(* IEC 61131-3 sources: SortJet_MasterSPS_Aufbau.fbsproj/07_Auftragsverwaltung/BasisSchrittketten (part 3) *)

(* ---- TS_Eintransport.fb.st ---- *)
(* METADATA
{
	"v3Meta": {
		"objectGuid": "2467a7d0-b543-4c0f-8e2f-d0f3bb8e773e"
	}
}
*)
FUNCTION_BLOCK TS_Eintransport
VAR_INPUT

  // BOOLEAN
  bpReset                : BOOL;

  // WORD
  wStation               : WORD;

  // STRUKTUR
  Auftragsdaten          : Auftragsdaten_ST;

END_VAR
VAR_OUTPUT

  // BOOLEAN
  bpDone                 : BOOL;
  bpFehler               : BOOL;

END_VAR
VAR
  // BOOLEAN
  blStationQuittiertScheiben : BOOL;

  // WORD
  wlEintransportstation  : WORD;

  // INT
  ilScheibenZuQuittieren : INT;

  // STEPS
  steplSchritt           : STEPS_TE;

END_VAR

//-------------------------------------------------------------------------------------------------
// STEUERUNG: EINTRANSPORT
//-------------------------------------------------------------------------------------------------
IF ( Auftragsdaten.wAuftrag = eStation_Eintransport ) THEN
  CASE steplSchritt OF
    // EINTRANSPORT  =============================== ============
    STEP_0_E:
      (* Hinweis:
         - Ueberpruefen des Sicherheitskreises
      *)
      IF  (checkSafetyCircuitsNotBlocked(starrTransferShuttleBasisParameter[wStation])
            AND NOT starrTransfershuttleBasisParameter[wStation].bReset )
      THEN
        steplSchritt := STEP_100_E;
      END_IF

    // EINTRANSPORT  ===========================================
    STEP_100_E:
      (* Anmerkung:
         - Zielstation abfragen ob diese bereit ist zum Austransport
      *)
      wlEintransportstation := Auftragsdaten.wTransferstationsNr1;
      ilScheibenZuQuittieren := WORD_TO_INT( Auftragsdaten.wAnzahlScheiben);

      CASE wlEintransportstation OF

          (* Hinweis:
             - Ruecktransport durch den Speicher beruecksichtigen
          *)
          cERSTES_INPUTSHUTTLE..cLETZTES_INPUTSHUTTLE,
            cERSTES_OUTPUTSHUTTLE..cLETZTES_OUTPUTSHUTTLE:
          IF ( Job_Shuttle.AuftragsdatenWand[Auftragsdaten.wTransferstationsNr1, Auftragsdaten.wTransferwand].wAuftrag = eStation_Austransport ) THEN
            steplSchritt := STEP_110_E;

          ELSE
            wpgFehlerdaten[0] := starrTransfershuttleBasisParameter[wStation].stMKs.stStationsNummern.NummerExtern;
            wpgFehlerdaten[1] := wlEintransportstation;
            wpgFehlerdaten[2] := Job_Shuttle.AuftragsdatenWand[Auftragsdaten.wTransferstationsNr1, Auftragsdaten.wTransferwand].wAuftrag;

            SpsError( eFehler_Station,
                      cMELDUNG_AUFTRAGSDATEN_AUFTRAGSTATUS_GLAS_SENDER_UNGUELTIG,
                      starrTransfershuttleBasisParameter[wStation].stMKs.stStationsNummern.NummerIntern,
                      AutomatikkreisBestimmen(starrTransfershuttleBasisParameter[wStation].stMKs.stStationsNummern.NummerSPS),
                      wpgFehlerdaten );

            steplSchritt := STEP_900_E;
          END_IF

        // Stationen
        //   - Wie beim Shuttle: Der TS legt den Austransport-Auftrag der Station an, sobald sie belegt ist
        cERSTE_STATION..cLETZTE_STATION:
          IF (    ( Job_Stationen.AuftragsdatenWand[wlEintransportstation, Auftragsdaten.wTransferwand].wAuftrag = eStation_Belegt )
               OR ( Job_Stationen.AuftragsdatenWand[wlEintransportstation, Auftragsdaten.wTransferwand].wAuftrag = eStation_Warte_Auf_Austransport ) )
             AND AutomatikAktiv(wlEintransportstation)
          THEN

            Job_Stationen.AuftragsdatenWand[wlEintransportstation, Auftragsdaten.wTransferwand]          := AuftragsdatenUmkopieren(FALSE, FALSE, Auftragsdaten);
            Job_Stationen.AuftragsdatenWand[wlEintransportstation, Auftragsdaten.wTransferwand].wAuftrag := eStation_Austransport;

            // Kopplung zur Station herstellen
            starrTransfershuttleBasisParameter[wStation].InGlasTransportNachfolger[cWAND_1] := starrStationBasisParameter[wlEintransportstation].OutGlasTransport[Auftragsdaten.wTransferwand];
            starrTransfershuttleBasisParameter[wStation].InGlasTransportVorgaenger[cWAND_1] := starrStationBasisParameter[wlEintransportstation].OutGlasTransport[Auftragsdaten.wTransferwand];

            steplSchritt := STEP_110_E;
          END_IF

        ELSE
          wpgFehlerdaten[0] := starrTransfershuttleBasisParameter[wStation].stMKs.stStationsNummern.NummerExtern;
          wpgFehlerdaten[1] := wlEintransportstation;

          SpsError( eFehler_Station,
                    cMELDUNG_AUFTRAGSDATEN_FALSCHE_EINLAUFSTATION,
                    starrTransfershuttleBasisParameter[wStation].stMKs.stStationsNummern.NummerIntern,
                    AutomatikkreisBestimmen(starrTransfershuttleBasisParameter[wStation].stMKs.stStationsNummern.NummerSPS),
                    wpgFehlerdaten );

          steplSchritt := STEP_900_E;

      END_CASE

      (* Fehlerbehandlung:
         - Shuttle
      *)
      IF ( starrTransfershuttleBasisParameter[wStation].bFehler ) THEN

        SpsError( eFehler_Station,
                  starrTransfershuttleBasisParameter[wStation].wFehlerNummer,
                  starrTransfershuttleBasisParameter[wStation].stMKs.stStationsNummern.NummerIntern,
                  AutomatikkreisBestimmen(starrTransfershuttleBasisParameter[wStation].stMKs.stStationsNummern.NummerSPS),
                  starrTransfershuttleBasisParameter[wStation].awFehlerInformationen );

        steplSchritt := STEP_900_E;
      END_IF

    // EINTRANSPORT  ===========================================
    STEP_110_E:

      (* Hinweis:
         - Starten des Eintransport
      *)
      IF ( Auftragsdaten.wTransferwand = cWAND_1 ) THEN
        starrTransfershuttleBasisParameter[wStation].bScheibentrennen[cWAND_1] := NOT Auftragsdaten.stAuftragsInformationen.cBIT_SRC_WALL_1_EMPTY;
      ELSE
        starrTransfershuttleBasisParameter[wStation].bScheibentrennen[cWAND_1] := NOT Auftragsdaten.stAuftragsInformationen.cBIT_SRC_WALL_2_EMPTY;
      END_IF

      starrTransfershuttleBasisParameter[wStation].pAuftrag[cWAND_1] := Auftragsdaten;
      starrTransfershuttleBasisParameter[wStation].bEintransport[cWAND_1] := TRUE;
      starrTransfershuttleBasisParameter[wStation].bRueckwaertsTransportieren[cWAND_1] := ( starrTransferShuttleBasisParameter[wStation].stMKs.stSchnittstellendaten.aEintransporte.Station[wlEintransportstation] = Rueckwaertig );

      steplSchritt := STEP_400_E;

    // EINTRANSPORT  ===========================================
    STEP_400_E:
      // ---------------------------------------------------------------------------------------
      //  QUITTIERUNGEN UND EINTRANSPORT- ABSCHLUSS
      //
      //  Hinweis:
      //  - Scheibenquittieren: Message zur MMI
      // ---------------------------------------------------------------------------------------

      IF ( starrTransfershuttleBasisParameter[wStation].OutGlasTransport[cWAND_1].bQuittScheibe ) THEN

        IF ( ilScheibenZuQuittieren > 0 ) AND starrTransfershuttleBasisParameter[wStation].stMKs.stSchnittstellendaten.aEintransporte.bStationQuittiertScheibe[wlEintransportstation] THEN

          wSps2MmiZielStation  := starrTransfershuttleBasisParameter[wStation].stMKs.stStationsNummern.NummerIntern;
          wSps2MmiQuellStation := Auftragsdaten.wTransferstationsNr1;
          wSps2MmiZielWand     := cWAND_1;
          wSps2MmiQuellWand    := Auftragsdaten.wTransferwand;
          dwSps2MmiWartezeit   := starrTransfershuttleBasisParameter[wStation].dwWartezeit[cWAND_1];
          wSPS2MMIAuftragstyp  := 0;

          MsgToMmi(auftragsnr_w := SB0_SPS_QUIT_SHEET_ORDER );
        END_IF

        ilScheibenZuQuittieren := ilScheibenZuQuittieren - 1;

      END_IF

      (* Hinweis:
         - Abschliessen des Eintransports ( Transfershuttle )
      *)
      IF( starrTransfershuttleBasisParameter[wStation].bEintransportAbgeschlossen[cWAND_1] ) THEN

        starrTransfershuttleBasisParameter[wStation].bEintransport[cWAND_1] := FALSE;
        steplSchritt := STEP_1000_E;

      END_IF

      (* Fehlerbehandlung:
         - Transfershuttle
      *)
      IF ( starrTransfershuttleBasisParameter[wStation].bFehler ) THEN

        IF ( aTransfershuttles[wStation].bpAnforderungBetriebsstopp ) THEN

          IF ( bgAktivierungTransfershuttleSystemcheck ) THEN
            wgSps2MmiShuttleNr                 := starrTransfershuttleBasisParameter[wStation].stMKs.stStationsNummern.NummerIntern;
            rgSPS2MMIExtractionShuttlePosition := starrTransfershuttleBasisParameter[wStation].rAktuellePositionQuerfahrt;
            wSps2MmiFehlertyp                  := aTransfershuttles[wStation].wpAusnahmefehlerTyp;
            MsgToMmi(auftragsnr_w := SB0_SPS_TRANSFERSHUTTLEFEHLER );// Fehlermeldung ans MMI für den folgenden Systemcheck
          END_IF

        END_IF

        starrTransfershuttleBasisParameter[wStation].bEintransport[cWAND_1] := FALSE;

        SpsError( eFehler_Station,
                  starrTransfershuttleBasisParameter[wStation].wFehlerNummer,
                  starrTransfershuttleBasisParameter[wStation].stMKs.stStationsNummern.NummerIntern,
                  AutomatikkreisBestimmen(starrTransfershuttleBasisParameter[wStation].stMKs.stStationsNummern.NummerSPS),
                  starrTransfershuttleBasisParameter[wStation].awFehlerInformationen );

        steplSchritt := STEP_900_E;

      END_IF

    // AUSTRANSPORT ==============================================
    STEP_410_E:
      (* Anmerkung:
         - Gueltige Anzahl von Scheiben wurden quittiert
      *)
      IF ( ilScheibenZuQuittieren = 0 ) THEN
        starrTransfershuttleBasisParameter[wStation].bEintransport[cWAND_1] := FALSE;
        steplSchritt := STEP_1000_E;

      (* Anmerkung:
         - Zu wenig Scheiben quittiert
      *)
      ELSIF ( ilScheibenZuQuittieren > 0 ) THEN
        wpgFehlerdaten[0] := starrTransfershuttleBasisParameter[wStation].stMKs.stStationsNummern.NummerExtern;
        wpgFehlerdaten[1] := cWAND_1;

        SpsError( eFehler_Station,
                  cMELDUNG_STATION_ZUWENIG_SCHEIBEN_QUITTIERT_WAND_EINTRANSPORT,
                  starrTransfershuttleBasisParameter[wStation].stMKs.stStationsNummern.NummerIntern,
                  AutomatikkreisBestimmen(starrTransfershuttleBasisParameter[wStation].stMKs.stStationsNummern.NummerSPS),
                  wpgFehlerdaten );

        starrTransfershuttleBasisParameter[wStation].bEintransport[cWAND_1] := FALSE;
        steplSchritt := STEP_900_E;

      (* Anmerkung:
         - Zu viele Scheiben quittiert
      *)
      ELSIF ( ilScheibenZuQuittieren < 0 ) THEN
        wpgFehlerdaten[0] := starrTransfershuttleBasisParameter[wStation].stMKs.stStationsNummern.NummerExtern;
        wpgFehlerdaten[1] := cWAND_1;

        SpsError( eFehler_Station,
                  cMELDUNG_STATION_ZUVIELE_SCHEIBEN_QUITTIERT_WAND_EINTRANSPORT,
                  starrTransfershuttleBasisParameter[wStation].stMKs.stStationsNummern.NummerIntern,
                  AutomatikkreisBestimmen(starrTransfershuttleBasisParameter[wStation].stMKs.stStationsNummern.NummerSPS),
                  wpgFehlerdaten );

        starrTransfershuttleBasisParameter[wStation].bEintransport[cWAND_1] := FALSE;
        steplSchritt := STEP_900_E;
      END_IF

    // EINTRANSPORT  ===========================================
    STEP_900_E:
      (* Hinweis:
         - Berücksichtigung wie Transportiert wurde
           => Wichtig: Automatikkreis beachten
      *)
      bpFehler := TRUE;

    // EINTRANSPORT  ===========================================
    STEP_1000_E:
      bpDone := TRUE;

      (* Hinweis:
         - Beenden des EIntransports [Bereit fuer den naechsten Auftrag]
      *)
      Auftragsdaten.wAuftrag := eStation_Kein_Auftrag;

      (* Hinweis:
         - Pruefen ob die Transferkopplung geloest werden muss
      *)
      IF ( PruefungWertImIntervall(Auftragsdaten.wTransferstationsNr2, cERSTES_TRANSFERSHUTTLE, cLETZTES_TRANSFERSHUTTLE) ) THEN

        IF ( Job_Shuttle.AuftragsdatenTransfershuttle[Auftragsdaten.wTransferstationsNr2].wAuftrag = eStation_Transportkopplung ) THEN
          Job_Shuttle.abpResetTransportkopplung[Auftragsdaten.wTransferstationsNr2] := TRUE;
        END_IF

      END_IF

  // EINTRANSPORT  ===========================================
  END_CASE
END_IF

IF bpReset THEN
  bpFehler := FALSE;
  bpDone := FALSE;
  bpReset := FALSE;
  starrTransfershuttleBasisParameter[wStation].bEintransport[cWAND_1] := FALSE;
  steplSchritt := STEP_0_E;
END_IF
END_FUNCTION_BLOCK

(* ---- TS_Querfahrt.fb.st ---- *)
(* METADATA
{
	"v3Meta": {
		"objectGuid": "302a3845-d7bd-4de5-be7f-afeb7baaa6cc"
	}
}
*)
FUNCTION_BLOCK TS_Querfahrt
VAR_INPUT

  // BOOLEAN
  bpReset                : BOOL;

  // WORD
  wStation               : WORD;

  // STRUKTUR
  Auftragsdaten          : Auftragsdaten_ST;

END_VAR
VAR_OUTPUT

  // BOOLEAN
  bpDone                 : BOOL;
  bpFehler               : BOOL;

END_VAR
VAR

  // STEPS
  steplSchritt           : STEPS_TE;

END_VAR

//-------------------------------------------------------------------------------------------------
// STEUERUNG: POSITIONIERUNG
//-------------------------------------------------------------------------------------------------
(* Hinweis [VERFAHRLOGIK]:
   - Das TS wird an eine mögliche neue Zielposition des nächsten echten Auftrages vorpositioniert,
     weil das dazugehörige Transfershuttle noch besetzt ist durch einen anderen Auftrag
*)
IF ( Auftragsdaten.wAuftrag = eStation_Vorabpositionierung) THEN

  CASE steplSchritt OF
    // POSITIONIERUNG ===========================================
    STEP_0_E:
      IF checkSafetyCircuitsNotBlocked(starrTransferShuttleBasisParameter[wStation])
         AND NOT starrTransfershuttleBasisParameter[wStation].bReset
      THEN

        IF ( ABS( starrTransfershuttleBasisParameter[wStation].rAktuellePositionQuerfahrt - Auftragsdaten.rVorabPosition ) <= rgMKZielPositionToleranz ) THEN
          steplSchritt := STEP_500_E;
        ELSIF starrTransfershuttleBasisParameter[wStation].stMKs.bDeaktivieren THEN
          steplSchritt := STEP_600_E;
        ELSE
          steplSchritt := STEP_10_E;
        END_IF

      END_IF

    // POSITIONIERUNG ===========================================
    STEP_10_E: // Positionere Shuttle
      (* Hinweis:
         - Uebergabe der Auftragsdaten
      *)
      starrTransfershuttleBasisParameter[wStation].pAuftragVorabPositionierung := Auftragsdaten;
      starrTransfershuttleBasisParameter[wStation].bVorabpositionieren := TRUE;

      steplSchritt := STEP_20_E;

    // POSITIONIERUNG ===========================================
    STEP_20_E:
      (* Hinweis:
         - Nachricht absetzen
      *)
      IF ( starrTransfershuttleBasisParameter[wStation].bUpdateVorabPositionieren = TRUE ) THEN

        wSps2MmiQuittVorabShuttleNr := starrTransfershuttleBasisParameter[wStation].stMKs.stStationsNummern.NummerIntern;
        rgSPS2MMIExtractionShuttlePosition := starrTransfershuttleBasisParameter[wStation].rAktuellePositionQuerfahrt;
        MsgToMmi(auftragsnr_w := SB0_SPS_SHUTTLEVORABPOSITIONIERUNGUPDATE );// Quit 2 MMI Scheibe vorne

        starrTransfershuttleBasisParameter[wStation].bUpdateVorabPositionieren := FALSE;

        steplSchritt := STEP_100_E;
      END_IF

      (* Fehlerbehandlung:
         - Inputshuttle
      *)
      IF ( starrTransfershuttleBasisParameter[wStation].bFehler ) THEN
        starrTransfershuttleBasisParameter[wStation].bVorabpositionieren := FALSE;

        SpsError( eFehler_Station,
                  starrTransfershuttleBasisParameter[wStation].wFehlerNummer,
                  starrTransfershuttleBasisParameter[wStation].stMKs.stStationsNummern.NummerIntern,
                  AutomatikkreisBestimmen(starrTransfershuttleBasisParameter[wStation].stMKs.stStationsNummern.NummerSPS),
                  starrTransfershuttleBasisParameter[wStation].awFehlerInformationen );

        steplSchritt := STEP_900_E;
      END_IF

    // POSITIONIERUNG ===========================================
    STEP_100_E:
      (* Hinweis:
         - Positionierung abgeschlossen
           => Nachricht absetzen
      *)
      IF NOT starrTransfershuttleBasisParameter[wStation].stMKs.bDeaktivieren THEN

        IF ( starrTransfershuttleBasisParameter[wStation].bVorabpositionierenAbgeschlossen ) THEN
          starrTransfershuttleBasisParameter[wStation].bVorabpositionieren := FALSE;

          wSps2MmiQuittVorabShuttleNr        := starrTransfershuttleBasisParameter[wStation].stMKs.stStationsNummern.NummerIntern;
          rgSPS2MMIExtractionShuttlePosition := aTransfershuttles[wStation].rpIstPositionNachPositionierung;
          MsgToMmi(auftragsnr_w := SB0_SPS_QUITTSHUTTLEVORABPOSITIONIERUNG );// Quit 2 MMI Scheibe vorne

          steplSchritt := STEP_1000_E;
        END_IF

      ELSE

        IF ( starrTransfershuttleBasisParameter[wStation].bVorabpositionierenAbgeschlossen ) THEN
          starrTransfershuttleBasisParameter[wStation].bVorabpositionieren := FALSE;

          wSps2MmiQuittVorabShuttleNr        := starrTransfershuttleBasisParameter[wStation].stMKs.stStationsNummern.NummerIntern;
          rgSPS2MMIExtractionShuttlePosition := Auftragsdaten.rVorabPosition;
          MsgToMmi(auftragsnr_w := SB0_SPS_QUITTSHUTTLEVORABPOSITIONIERUNG );// Quit 2 MMI Scheibe vorne

          steplSchritt := STEP_1000_E;
        END_IF

      END_IF

      (* Fehlerbehandlung:
         - Inputshuttle
      *)
      IF ( starrTransfershuttleBasisParameter[wStation].bFehler ) THEN
        starrTransfershuttleBasisParameter[wStation].bVorabpositionieren := FALSE;

        SpsError( eFehler_Station,
                  starrTransfershuttleBasisParameter[wStation].wFehlerNummer,
                  starrTransfershuttleBasisParameter[wStation].stMKs.stStationsNummern.NummerIntern,
                  AutomatikkreisBestimmen(starrTransfershuttleBasisParameter[wStation].stMKs.stStationsNummern.NummerSPS),
                  starrTransfershuttleBasisParameter[wStation].awFehlerInformationen );

        steplSchritt := STEP_900_E;
      END_IF

    // POSITIONIERUNG ===========================================
    STEP_500_E:
      wSps2MmiQuittVorabShuttleNr := starrTransfershuttleBasisParameter[wStation].stMKs.stStationsNummern.NummerIntern;
      rgSPS2MMIExtractionShuttlePosition := starrTransfershuttleBasisParameter[wStation].rAktuellePositionQuerfahrt;
      MsgToMmi(auftragsnr_w := SB0_SPS_SHUTTLEVORABPOSITIONIERUNGUPDATE );// Quit 2 MMI Scheibe vorne
      steplSchritt := STEP_510_E;

    // POSITIONIERUNG ===========================================
    STEP_510_E:
      wSps2MmiQuittVorabShuttleNr        := starrTransfershuttleBasisParameter[wStation].stMKs.stStationsNummern.NummerIntern;
      rgSPS2MMIExtractionShuttlePosition := starrTransfershuttleBasisParameter[wStation].rAktuellePositionQuerfahrt;
      MsgToMmi(auftragsnr_w := SB0_SPS_QUITTSHUTTLEVORABPOSITIONIERUNG );// Quit 2 MMI Scheibe vorne
      steplSchritt := STEP_1000_E;

    // POSITIONIERUNG ===========================================
    STEP_600_E:
      wSps2MmiQuittVorabShuttleNr := starrTransfershuttleBasisParameter[wStation].stMKs.stStationsNummern.NummerIntern;
      rgSPS2MMIExtractionShuttlePosition := Auftragsdaten.rVorabPosition;
      MsgToMmi(auftragsnr_w := SB0_SPS_SHUTTLEVORABPOSITIONIERUNGUPDATE );// Quit 2 MMI Scheibe vorne
      steplSchritt := STEP_610_E;

    // POSITIONIERUNG ===========================================
    STEP_610_E:
      wSps2MmiQuittVorabShuttleNr        := starrTransfershuttleBasisParameter[wStation].stMKs.stStationsNummern.NummerIntern;
      rgSPS2MMIExtractionShuttlePosition := Auftragsdaten.rVorabPosition;
      MsgToMmi(auftragsnr_w := SB0_SPS_QUITTSHUTTLEVORABPOSITIONIERUNG );// Quit 2 MMI Scheibe vorne
      steplSchritt := STEP_1000_E;

    // POSITIONIERUNG ===========================================
    STEP_900_E:
      bpFehler := TRUE;

    // POSITIONIERUNG ===========================================
    STEP_1000_E:
      bpDone := TRUE;
      Auftragsdaten.wAuftrag := eStation_Kein_Auftrag;

  // POSITIONIERUNG ===========================================
  END_CASE

END_IF

IF bpReset THEN
  bpFehler := FALSE;
  bpDone := FALSE;
  bpReset := FALSE;
  starrTransfershuttleBasisParameter[wStation].bUpdateVorabPositionieren := FALSE;
  starrTransfershuttleBasisParameter[wStation].bVorabpositionieren := FALSE;
  steplSchritt := STEP_0_E;
END_IF
END_FUNCTION_BLOCK

(* ---- TS_Transportkopplung.fb.st ---- *)
(* METADATA
{
	"v3Meta": {
		"objectGuid": "b272f643-831b-42e0-8c4f-868bd25374f4"
	}
}
*)
FUNCTION_BLOCK TS_Transportkopplung
VAR_INPUT

  // BOOLEAN
  bpReset                : BOOL;

  // WORD
  wStation               : WORD;

  // STRUKTUR
  Auftragsdaten          : Auftragsdaten_ST;

END_VAR
VAR_OUTPUT

  // BOOLEAN
  bpDone                 : BOOL;
  bpFehler               : BOOL;

END_VAR
VAR

  // STEPS
  steplSchritt           : STEPS_TE;

END_VAR
//-------------------------------------------------------------------------------------------------
// STEUERUNG: TRANSPORTKOPPLUNG
//-------------------------------------------------------------------------------------------------
IF ( Auftragsdaten.wAuftrag = eStation_Transportkopplung ) THEN
  CASE steplSchritt OF
    // TRANSPORTKOPPLUNG ===========================================
    STEP_0_E:
      (* Hinweis:
         - Ueberpruefen des Sicherheitskreises
      *)
      IF checkSafetyCircuitsNotBlocked(starrStationBasisParameter[wStation])
         AND NOT starrTransfershuttleBasisParameter[wStation].bReset
      THEN
        steplSchritt := STEP_100_E;
      END_IF

    // TRANSPORTKOPPLUNG ===========================================
    STEP_100_E:

      starrTransfershuttleBasisParameter[wStation].pAuftrag[cWAND_1] := Auftragsdaten;
      starrTransfershuttleBasisParameter[wStation].bTransportkopplung[cWAND_1] := TRUE;

      steplSchritt := STEP_110_E;

    // TRANSPORTKOPPLUNG ===========================================
    STEP_110_E:
      (* Fehlerbehandlung:
         - Transfershuttle
      *)
      IF ( starrTransfershuttleBasisParameter[wStation].bFehler ) THEN

        starrTransfershuttleBasisParameter[wStation].bTransportkopplung[cWAND_1] := FALSE;

        SpsError( eFehler_Station,
                  starrTransfershuttleBasisParameter[wStation].wFehlerNummer,
                  starrTransfershuttleBasisParameter[wStation].stMKs.stStationsNummern.NummerIntern,
                  AutomatikkreisBestimmen(starrTransfershuttleBasisParameter[wStation].stMKs.stStationsNummern.NummerSPS),
                  starrTransfershuttleBasisParameter[wStation].awFehlerInformationen );

        steplSchritt := STEP_900_E;

      END_IF

    // TRANSPORTKOPPLUNG ===========================================
    STEP_900_E:
      bpFehler := TRUE;

    // TRANSPORTKOPPLUNG ===========================================
    STEP_1000_E:
      bpDone := TRUE;

  // TRANSPORTKOPPLUNG ===========================================
  END_CASE
END_IF

IF bpReset THEN
  starrTransfershuttleBasisParameter[wStation].bTransportkopplung[cWAND_1] := FALSE;
  steplSchritt := STEP_0_E;
  bpFehler := FALSE;
  bpDone := FALSE;
  bpReset := FALSE;
END_IF
END_FUNCTION_BLOCK

(* ---- TS_Vortransport.fb.st ---- *)
(* METADATA
{
	"v3Meta": {
		"objectGuid": "82a7ab83-6d97-4992-8583-d2407cc9730b"
	}
}
*)
FUNCTION_BLOCK TS_Vortransport
VAR_INPUT

  // BOOLEAN
  bpReset                : BOOL;

  // WORD
  wStation               : WORD;

  // STRUKTUR
  Auftragsdaten          : Auftragsdaten_ST;

END_VAR
VAR_OUTPUT

  // BOOLEAN
  bpDone                 : BOOL;
  bpFehler               : BOOL;

END_VAR
VAR

  // WORD
  wlVerbundStation       : WORD;

  // STEPS
  steplSchritt           : STEPS_TE;

END_VAR
//-------------------------------------------------------------------------------------------------
// STEUERUNG: VORTRANSPORT
//-------------------------------------------------------------------------------------------------
IF ( Auftragsdaten.wAuftrag = eStation_Vortransport ) THEN
  CASE steplSchritt OF
    // VORTRANSPORT ==============================================
    STEP_0_E:
      IF (  checkSafetyCircuitsNotBlocked(starrStationBasisParameter[wStation])
           AND NOT starrTransfershuttleBasisParameter[wStation].bReset )
      THEN

        steplSchritt := STEP_100_E;

        IF ( Auftragsdaten.rStationsZielposition > aTransfershuttles[wStation].Querfahrt.Antrieb.rpMaxPosition ) THEN
          wpgFehlerdaten[0] := wStation;
          SysMemCpy( ADR( wpgFehlerdaten[1] ), ADR ( aTransfershuttles[wStation].Querfahrt.Antrieb.rpMaxPosition ), 4 );
          SysMemCpy( ADR( wpgFehlerdaten[3] ), ADR ( Auftragsdaten.rStationsZielposition ), 4 );

          SpsError( eFehler_Station,
                    cMELDUNG_AUFTRAGSDATEN_ZIELPOSITION_ZU_GROSS,
                    starrTransfershuttleBasisParameter[wStation].stMKs.stStationsNummern.NummerIntern,
                    AutomatikkreisBestimmen(starrTransfershuttleBasisParameter[wStation].stMKs.stStationsNummern.NummerSPS),
                    wpgFehlerdaten );

          steplSchritt := STEP_900_E;
        END_IF

        IF ( Auftragsdaten.rStationsZielposition < aTransfershuttles[wStation].Querfahrt.Antrieb.rpMinPosition ) THEN
          wpgFehlerdaten[0] := wStation;
          SysMemCpy( ADR( wpgFehlerdaten[1] ), ADR ( aTransfershuttles[wStation].Querfahrt.Antrieb.rpMinPosition ), 4 );
          SysMemCpy( ADR( wpgFehlerdaten[3] ), ADR ( Auftragsdaten.rStationsZielposition ), 4 );

          SpsError( eFehler_Station,
                    cMELDUNG_AUFTRAGSDATEN_ZIELPOSITION_ZU_KLEIN,
                    starrTransfershuttleBasisParameter[wStation].stMKs.stStationsNummern.NummerIntern,
                    AutomatikkreisBestimmen(starrTransfershuttleBasisParameter[wStation].stMKs.stStationsNummern.NummerSPS),
                    wpgFehlerdaten );
          steplSchritt := STEP_900_E;
        END_IF

      END_IF

    // VORTRANSPORT ==============================================
    STEP_100_E:
      // ---------------------------------------------------------------------------------------
      //  PRUEFEN TRANSFERSHUTTLE VERBUND
      //
      //  Hinweis:
      //  - Transferstation2 = 0   => Vortransport mit nur einem Transfershuttle
      //  - Transferstation2 <> 0  => Vortransport im Transfershuttle-Verbund
      // ---------------------------------------------------------------------------------------

      IF ( Auftragsdaten.wTransferstationsNr2 = 0 ) THEN

        IF ( NOT starrTransfershuttleBasisParameter[wStation].bAuftragAktiv ) THEN
          starrTransfershuttleBasisParameter[wStation].pAuftrag[cWAND_1]      := Auftragsdaten;
          aTransfershuttles[wStation].rpVorpositionierWeg                     := Auftragsdaten.rAuftragsLaenge;
          starrTransfershuttleBasisParameter[wStation].bVortransport[cWAND_1] := TRUE;
          steplSchritt := STEP_400_E;
        END_IF

      ELSE
        wlVerbundStation := Auftragsdaten.wTransferstationsNr2;

        IF ( Job_Shuttle.AuftragsdatenTransfershuttle[Auftragsdaten.wTransferstationsNr2].wAuftrag = eStation_Kein_Auftrag ) THEN
          steplSchritt := STEP_200_E;
        END_IF

      END_IF

    // VORTRANSPORT ==============================================
    STEP_200_E:
      // ---------------------------------------------------------------------------------------
      //  TRANSFERSHUTTLE VERBUND
      //
      //  Hinweis:
      //  - n/c
      // ---------------------------------------------------------------------------------------

      IF ( NOT starrTransfershuttleBasisParameter[wStation].bAuftragAktiv ) THEN

        (* Hinweis:
           - Transfershuttle koppeln
        *)
        aTransfershuttles[wStation].stpInTransportVerbund                             := aTransfershuttles[wlVerbundStation].stpOutTransportVerbund;
        aTransfershuttles[wlVerbundStation].stpInTransportVerbund  := aTransfershuttles[wStation].stpOutTransportVerbund;

        (* Hinweis:
           - Auftragsdaten uebergeben
        *)
        Job_Shuttle.AuftragsdatenTransfershuttle[wlVerbundStation].rStationsZielposition := Auftragsdaten.rTransferposition2 ;
        Job_Shuttle.AuftragsdatenTransfershuttle[wlVerbundStation].wStationsNr           := Auftragsdaten.wTransferstationsNr2 ;
        Job_Shuttle.AuftragsdatenTransfershuttle[wlVerbundStation].wAuftrag:= eStation_Transportkopplung;

        (* Hinweis:
           - Auftragsdaten uebergeben
        *)
        starrTransfershuttleBasisParameter[wStation].pAuftrag[cWAND_1]      := Auftragsdaten;
        aTransfershuttles[wStation].rpVorpositionierWeg                     := Auftragsdaten.rAuftragsLaenge;
        starrTransfershuttleBasisParameter[wStation].bVortransport[cWAND_1] := TRUE;

        steplSchritt := STEP_400_E;

      END_IF

    // VORTRANSPORT ==============================================
    STEP_400_E:
      // ---------------------------------------------------------------------------------------
      //  TRANSFERSHUTTLE VORTRANSPORT ABGESCHLOSSEN
      //
      //  Hinweis:
      //  - n/c
      // ---------------------------------------------------------------------------------------

      IF ( starrTransfershuttleBasisParameter[wStation].bVortransportAbgeschlossen[cWAND_1] ) THEN

        (* Hinweis:
           - Nachricht an die HMMI
        *)
        wSps2MmiQuittierungVortransportStationsNr1 := starrTransfershuttleBasisParameter[wStation].stMKs.stStationsNummern.NummerIntern;
        wSps2MmiQuittierungVortransportStationsNr2 := Auftragsdaten.wTransferstationsNr2;
        wSps2MmiQuittierungVortransportStatus      := 1; // 0  = nicht Erfolgreich / 1 = erfolgreich
        rSps2MmiQuittierungVortransportWegStrecke  := aTransfershuttles[wStation].rpVorpositionierterWeg;

        MsgToMmi(auftragsnr_w := SB0_SPS_SortierungQuittExtractionShuttleData );

        starrTransfershuttleBasisParameter[wStation].bVortransport[cWAND_1] := FALSE;

        steplSchritt := STEP_1000_E;
      END_IF

      (* Hinweis:
         - -Ausnahmefehler
      *)
      IF ( starrTransfershuttleBasisParameter[wStation].bFehler ) THEN
        SpsError( eFehler_Station,
                  starrTransfershuttleBasisParameter[wStation].wFehlerNummer,
                  starrTransfershuttleBasisParameter[wStation].stMKs.stStationsNummern.NummerIntern,
                  AutomatikkreisBestimmen(starrTransfershuttleBasisParameter[wStation].stMKs.stStationsNummern.NummerSPS),
                  starrTransfershuttleBasisParameter[wStation].awFehlerInformationen );

        starrTransfershuttleBasisParameter[wStation].bVortransport[cWAND_1] := FALSE;

        steplSchritt := STEP_900_E;
      END_IF

    // VORTRANSPORT ==============================================
    STEP_900_E:
      bpFehler := TRUE;

    // VORTRANSPORT ==============================================
    STEP_1000_E:
      bpDone := TRUE;

      Auftragsdaten.wAuftrag := eStation_Kein_Auftrag;

      (* Hinweis:
         - Pruefen ob die Transferkopplung geloest werden muss
      *)
      IF ( PruefungWertImIntervall(Auftragsdaten.wTransferstationsNr2, cERSTES_TRANSFERSHUTTLE, cLETZTES_TRANSFERSHUTTLE) ) THEN

        IF ( Job_Shuttle.AuftragsdatenTransfershuttle[Auftragsdaten.wTransferstationsNr2].wAuftrag = eStation_Transportkopplung ) THEN
          Job_Shuttle.AuftragsdatenTransfershuttle[Auftragsdaten.wTransferstationsNr2].wAuftrag := eStation_Kein_Auftrag;
        END_IF

      END_IF

  // VORTRANSPORT ==============================================
  END_CASE
END_IF

IF bpReset THEN
  starrTransfershuttleBasisParameter[wStation].bVortransport[cWAND_1] := FALSE;
  bpDone   := FALSE;
  bpReset  := FALSE;
  bpFehler := FALSE;
  steplSchritt := STEP_0_E;
END_IF
END_FUNCTION_BLOCK
